(* IEC 61131-3 sources: PLC-Static-Analysis/modules/plc-rules/src/test/resources/PLCA-Q006, 2 files *)

(* ---- compliant.st ---- *)
FUNCTION_BLOCK FB_InOk
VAR_INPUT
    bIn : BOOL;
    pIn : POINTER TO INT;
    refIn : REFERENCE TO INT;
END_VAR
VAR_IN_OUT
    nInOut : INT;
END_VAR
VAR
    bCopy : BOOL;
END_VAR
bCopy := bIn;
pIn^ := 1;
refIn := 2;
nInOut := 3;
END_FUNCTION_BLOCK

PROGRAM P_Caller
VAR
    fb : FB_InOk;
    n : INT;
END_VAR
fb.bIn := TRUE;
fb(bIn := FALSE, nInOut := n);
END_PROGRAM

(* ---- noncompliant.st ---- *)
TYPE ST_Pt :
STRUCT
    x : INT;
    y : INT;
END_STRUCT
END_TYPE

FUNCTION_BLOCK FB_In
VAR_INPUT
    bIn : BOOL;
    nIn : INT;
    stIn : ST_Pt;
END_VAR
bIn := FALSE; // PLCA-Q006
stIn.x := 0; // PLCA-Q006

METHOD M
VAR_INPUT
    nArg : INT;
END_VAR
nIn := 5; // PLCA-Q006
nArg := 0; // PLCA-Q006
END_METHOD
END_FUNCTION_BLOCK

FUNCTION_BLOCK FB_In2 EXTENDS FB_In
nIn := 1; // PLCA-Q006
END_FUNCTION_BLOCK

FUNCTION F_In : INT
VAR_INPUT
    n : INT;
END_VAR
n := n + 1; // PLCA-Q006
F_In := n;
END_FUNCTION
